Staubli VAL3: cycle_start.pgx

public program cycle_start()
begin
  rs:bToStartCycle=true
  wait(rs:bIsCycle==true)
  rs:bToStartCycle=false


  logMsg("PLC:startcycle")
end
